Universal Robots URScript: Prog_Name_That_Is_Very_Long_123.script

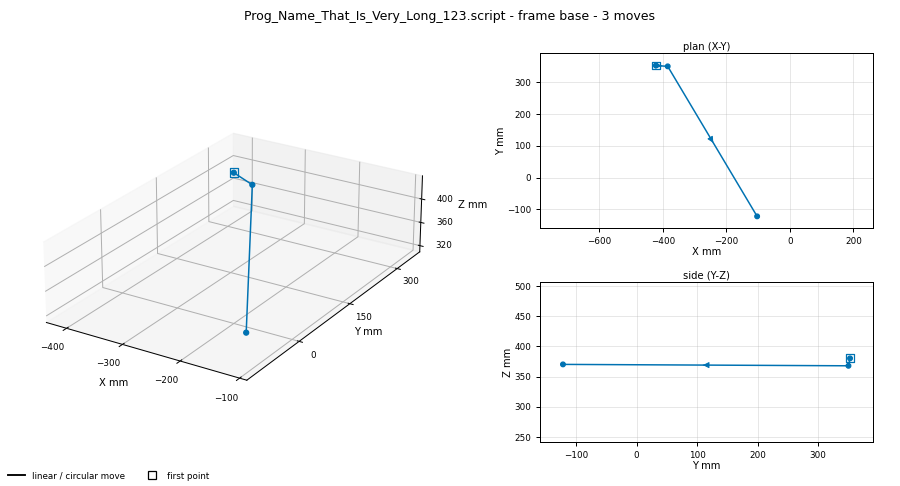
[picture p0: tool path of Prog_Name_That_Is_Very_Long_123.script in frame base, 3 of 5 moves have a stored position in this frame; points joined in program order, loops and branches not executed]
def Prog_Name_That_Is_Very_Long_123():
  # Global parameters:
  global speed_ms    = 0.250
  global speed_rads  = 0.750
  global accel_mss   = 1.200
  global accel_radss = 1.200
  global blend_radius_m = 0.000

  #--------------------------
  # Add any default subprograms here
  # For example, to drive a gripper as a program call:
  # def Gripper_Open():
  #   ...
  # end
  #
  # Example to drive a spray gun:
  def SprayOn(value):
    # use the value as an output:
    DO_SPRAY = 5
    if value == 0:
      set_standard_digital_out(DO_SPRAY, False)
    else:
      set_standard_digital_out(DO_SPRAY, True)
    end
  end

  # Example to synchronize 2
  def Synchronize():
    # Use the following digital output to signal the state of the robot:
    DO_SYNC = 1

    # Use the following digital input to get the state of another robot:
    DI_SYNC = 1

    if (get_standard_digital_out(DO_SYNC) == get_standard_digital_in(DI_SYNC)):
      set_standard_digital_out(DO_SYNC, not (get_standard_digital_out(DI_SYNC)))
      sleep(0.1)
      thread Thread_wait_1():
        while (True):
          sleep(0.01)
        end
      end
      if (get_standard_digital_out(DO_SYNC) != get_standard_digital_in(DI_SYNC)):
        global thread_handler_1=run Thread_wait_1()
        while (get_standard_digital_out(DO_SYNC) != get_standard_digital_in(DI_SYNC)):
          sync()
        end
        kill thread_handler_1
      end
    else:
      if (get_standard_digital_out(DO_SYNC) != get_standard_digital_in(DI_SYNC)):
        set_standard_digital_out(DO_SYNC, not (get_standard_digital_out(DO_SYNC)))
      end
    end
  end

  #
  # Example to move an external axis
  def MoveAxis(value):
    # use the value as an output:
    DO_AXIS_1 = 1
    DI_AXIS_1 = 1
    if value <= 0:
      set_standard_digital_out(DO_AXIS_1, False)

      # Wait for digital input to change state
      #while (get_standard_digital_in(DI_AXIS_1) != False):
      #  sync()
      #end
    else:
      set_standard_digital_out(DO_AXIS_1, True)

      # Wait for digital input to change state
      #while (get_standard_digital_in(DI_AXIS_1) != True):
      #  sync()
      #end
    end
  end
  #--------------------------


  # Main program:
  # Program generated by VerticalBot Studio for UR5e on 25/10/2026 12:00:00
  # Using nominal kinematics.
  # Using Ref. UR5e Base: p[0.000000, 0.000000, 0.000000, 0.000000, 0.000000, 0.000000]
  # set_reference(p[0.000000, 0.000000, 0.000000, 0.000000, 0.000000, 0.000000])
  # Using TCP Spindle: p[0.010000, 0.000000, 0.120000, 0.000000, 0.261799, 0.000000]
  set_tcp(p[0.010000, 0.000000, 0.120000, 0.000000, 0.261799, 0.000000])
  speed_ms    = 1.0000
  blend_radius_m = 0.0100
  movej([-0.523599, -1.745329, 1.570796, -1.396263, -1.570796, 0.349066],1.20000,0.75000,0,0.0000)
  movel(p[-0.421760, 0.353029, 0.380392, 3.048452, 0.496356, 0.454618],accel_mss,speed_ms,0,0.010)
  blend_radius_m = 0.0005
  movel(p[-0.384494, 0.350433, 0.368074, 3.036811, 0.389569, 0.461666],accel_mss,speed_ms,0,0.001)
  halt() # reimplement this function to force stop
  sleep(1.500)
  popup("Say "hi" to the operator","Message",False,False,blocking=False)
  # A long comment line that exceeds the usual controller limits for comments by far, really
  set_standard_digital_out(12, False)
  OUT_A = True
  while (get_standard_digital_in(4) != False):
    sync()
  end
  while (IN_B != True):
    sync()
  end
  Program_With_A_Long_Name_ABCDEFGHIJ()
  # Using Ref. Frame 12: p[0.250000, 0.300000, -0.010000, 0.000000, 0.000000, 1.570796]
  # set_reference(p[0.250000, 0.300000, -0.010000, 0.000000, 0.000000, 1.570796])
  # Using TCP Tool 7: p[0.010000, 0.000000, 0.120000, 0.000000, 0.261799, 0.000000]
  set_tcp(p[0.010000, 0.000000, 0.120000, 0.000000, 0.261799, 0.000000])
  speed_rads  = 0.5236
  accel_radss = 1.745
  movel(p[-0.103029, -0.121760, 0.370392, -1.712677, -2.378873, -0.325743],accel_mss,speed_ms,0,0.001)
  blend_radius_m = 0.0000
  movej([-0.523599, -1.745329, 1.570796, -1.396263, -1.570796, 0.349066],1.74533,0.52360,0,0.0000)
  # End of main program
end

Prog_Name_That_Is_Very_Long_123()
